TYPE ST_MAIN_VIS :
STRUCT
  eInitXts          : E_PROGRESS;
  sInitXts          : STRING(20);

  eInitApplication  : E_PROGRESS;
  sInitApplication  : STRING(20);

  nStateApplication : UINT;
END_STRUCT
END_TYPE

(* stored: Version 1.1.0.1
   DUT ST_MAIN_VIS: Id {863e53a0-0be7-4ab3-b120-ada52aee8a57} *)
